Fanuc KAREL source: IO0207.KL

PROGRAM IO0207
%NOLOCKGROUP
ROUTINE RTEST
VAR
L1 : ARRAY[3] OF INTEGER;L2 : XYZWPR
L3 : JOINTPOS9
L4 : POSITION
S1:INTEGER
S2:INTEGER
A:REAL
B:BOOLEAN
C:REAL
BEGIN
--
--
S1=1
L1[1]=2
B=TRUE
C=1.0
SET_INT_REG(S1,S1,S2)
END RTEST
BEGIN
RTEST
END IO0207
